FUNCTION FC 1 : VOID
BEGIN
NETWORK
      L P#M0.0
END_FUNCTION
